TYPE ST_BmsProt :
STRUCT
	eBatAction	: E_BatAction;		// 이 BMS에 걸린 가장 센 조치
	nModule		: UINT;				// 조치를 건 보호 모듈 ID
END_STRUCT
END_TYPE

(* stored: Version 1.1.0.1, ProductVersion 3.1.4024.15
   DUT ST_BmsProt: Id {8f52c4e2-3df1-4948-8829-c01546796ad8} *)
